                                   //LCom Version V1
                                   #statSend.tsendFct.data[#statSend.tsendFct.dataOffset] := #statSend.configTelegramV1.LComVersion;
                                   #statSend.tsendFct.data[#statSend.tsendFct.dataOffset + 1] := 16#03;
                                   #statSend.tsendFct.data[#statSend.tsendFct.dataOffset + 2] := #statSend.configTelegramV1.comMode;//ComMode
                                   #statSend.tsendFct.data[#statSend.tsendFct.dataOffset + 3] := #statSend.configTelegramV1.slidingWindow;//SlidingWindow
                                   //cycleTime
                                   #statSend.tsendFct.data[#statSend.tsendFct.dataOffset + 4] := #statSend.configTelegramV1.cycleTime.%B1;
                                   #statSend.tsendFct.data[#statSend.tsendFct.dataOffset + 5] := #statSend.configTelegramV1.cycleTime.%B0;
                                   //ackTimeOut
                                   #statSend.tsendFct.data[#statSend.tsendFct.dataOffset + 6] := #statSend.configTelegramV1.ackTimeOut.%B1;
                                   #statSend.tsendFct.data[#statSend.tsendFct.dataOffset + 7] := #statSend.configTelegramV1.ackTimeOut.%B0;
                                   //lifeSignCycle
                                   #statSend.tsendFct.data[#statSend.tsendFct.dataOffset + 8] := #statSend.configTelegramV1.lifeSignCycle.%B1;
                                   #statSend.tsendFct.data[#statSend.tsendFct.dataOffset + 9] := #statSend.configTelegramV1.lifeSignCycle.%B0;
                                   //status
                                   #statSend.tsendFct.data[#statSend.tsendFct.dataOffset + 10] := #statSend.configTelegramV1.status;
                                   //sendModeSyncTime
                                   #statSend.tsendFct.data[#statSend.tsendFct.dataOffset + 11] := #statSend.configTelegramV1.sendModeSyncTime;
                                   //maxSendDataLength
                                   #statSend.tsendFct.data[#statSend.tsendFct.dataOffset + 12] := #statSend.configTelegramV1.maxSendDataLength.%B1;
                                   #statSend.tsendFct.data[#statSend.tsendFct.dataOffset + 13] := #statSend.configTelegramV1.maxSendDataLength.%B0;
                                   //maxReceiveDataLength
                                   #statSend.tsendFct.data[#statSend.tsendFct.dataOffset + 14] := #statSend.configTelegramV1.maxReceiveDataLength.%B1;
                                   #statSend.tsendFct.data[#statSend.tsendFct.dataOffset + 15] := #statSend.configTelegramV1.maxReceiveDataLength.%B0;
                                   //calculate new offset
                                   #statSend.tsendFct.dataOffset := 16;
                               ELSE
                                   #statSend.tsendFct.data[#statSend.tsendFct.dataOffset] := #statSend.configTelegramV2.LComVersion;
                                   #statSend.tsendFct.data[#statSend.tsendFct.dataOffset + 1] := 16#03;
                                   //status
                                   #statSend.tsendFct.data[#statSend.tsendFct.dataOffset + 2] := #statSend.configTelegramV2.status;
                                   //sendModeSyncTime
                                   #statSend.tsendFct.data[#statSend.tsendFct.dataOffset + 3] := #statSend.configTelegramV2.sendModeSyncTime;
                                   //lifeSignCycle
                                   #tempDWord := TIME_TO_DWORD(#statSend.configTelegramV2.lifeSignCycle);
                                   #statSend.tsendFct.data[#statSend.tsendFct.dataOffset + 4] := #tempDWord.%B3;
                                   #statSend.tsendFct.data[#statSend.tsendFct.dataOffset + 5] := #tempDWord.%B2;
                                   #statSend.tsendFct.data[#statSend.tsendFct.dataOffset + 6] := #tempDWord.%B1;
                                   #statSend.tsendFct.data[#statSend.tsendFct.dataOffset + 7] := #tempDWord.%B0;
                                   //cycleTime
                                   #tempDWord := TIME_TO_DWORD(#statSend.configTelegramV2.cycleTime);
                                   #statSend.tsendFct.data[#statSend.tsendFct.dataOffset + 8] := #tempDWord.%B3;
                                   #statSend.tsendFct.data[#statSend.tsendFct.dataOffset + 9] := #tempDWord.%B2;
                                   #statSend.tsendFct.data[#statSend.tsendFct.dataOffset + 10] := #tempDWord.%B1;
                                   #statSend.tsendFct.data[#statSend.tsendFct.dataOffset + 11] := #tempDWord.%B0;
                                   //ackTimeOut
                                   #tempDWord := TIME_TO_DWORD(#statSend.configTelegramV2.ackTimeOut);
                                   #statSend.tsendFct.data[#statSend.tsendFct.dataOffset + 12] := #tempDWord.%B3;
                                   #statSend.tsendFct.data[#statSend.tsendFct.dataOffset + 13] := #tempDWord.%B2;
                                   #statSend.tsendFct.data[#statSend.tsendFct.dataOffset + 14] := #tempDWord.%B1;
                                   #statSend.tsendFct.data[#statSend.tsendFct.dataOffset + 15] := #tempDWord.%B0;
                                   //maxSendDataLength
                                   #statSend.tsendFct.data[#statSend.tsendFct.dataOffset + 16] := #statSend.configTelegramV2.maxSendDataLength.%B3;
                                   #statSend.tsendFct.data[#statSend.tsendFct.dataOffset + 17] := #statSend.configTelegramV2.maxSendDataLength.%B2;
                                   #statSend.tsendFct.data[#statSend.tsendFct.dataOffset + 18] := #statSend.configTelegramV2.maxSendDataLength.%B1;
                                   #statSend.tsendFct.data[#statSend.tsendFct.dataOffset + 19] := #statSend.configTelegramV2.maxSendDataLength.%B0;
                                   //maxReceiveDataLength
                                   #statSend.tsendFct.data[#statSend.tsendFct.dataOffset + 20] := #statSend.configTelegramV2.maxReceiveDataLength.%B3;
                                   #statSend.tsendFct.data[#statSend.tsendFct.dataOffset + 21] := #statSend.configTelegramV2.maxReceiveDataLength.%B2;
                                   #statSend.tsendFct.data[#statSend.tsendFct.dataOffset + 22] := #statSend.configTelegramV2.maxReceiveDataLength.%B1;
                                   #statSend.tsendFct.data[#statSend.tsendFct.dataOffset + 23] := #statSend.configTelegramV2.maxReceiveDataLength.%B0;
                                   //calculate new offset
                                   #statSend.tsendFct.dataOffset := 24;
                               END_IF;
                               #statSend.tsendFct.enable := TRUE;

                               #instLocalLifeSignCycleTimer(IN := FALSE,
                                                            PT := #diagnostics.localConfig.connection.lifeSignCycleTime);
                           ELSE
                               ;//Telegram 3 don´t need be send

                           END_IF;
                       ELSIF (NOT #diagnostics.localConfig.connection.useLComProtocol //without LCom Protocol
                           AND #statState.sender = #STATE_INACTIVE) THEN
                           #statSend.tsendFct.enable := FALSE;
                       ELSE
                           #statSend.tsendFct.enable := TRUE;

                           #instLocalLifeSignCycleTimer(IN := FALSE,
                                                        PT := #diagnostics.localConfig.connection.lifeSignCycleTime);
                       END_IF;

                       //differ between different connection types (IPv4, QDN)
                       IF (#diagnostics.localConfig.connection.connectType = #CON_TYPE_IPV4) THEN
                           #tempConnOucId := #statTconPar.ID;
                       ELSE    //#CON_TYPE_QDN
                           #tempConnOucId := #statTconParQdn.ID;
                       END_IF;

                       #instTSEND(REQ := #statSend.tsendFct.enable,
                                  LEN := #statSend.tsendFct.dataOffset,
                                  ID := #tempConnOucId,
                                  DATA := #statSend.tsendFct.data,
                                  STATUS => #statSend.tsendFct.status);

                       //16#80C4=Temporary communication error
                       IF (#statSend.tsendFct.status = 16#80C4) THEN

                           #instSendErrorTimer(IN := TRUE,
                                               PT := #MAX_TRIAL_TIME);

                           //#MAX_TRIAL_TIME is expired
                           IF #instSendErrorTimer.Q THEN
                               //Write diagnostics
                               #statDiag.bufferIndex := #statDiag.bufferIndex + 1;
                               #statDiag.buffer[#statDiag.bufferIndex].status := #ERR_SEND;
                               #statDiag.buffer[#statDiag.bufferIndex].subFunctionErrorID := #statSend.tsendFct.status;
                               #statDiag.buffer[#statDiag.bufferIndex].additionalValue1 := 0.0;
                               #statDiag.buffer[#statDiag.bufferIndex].additionalValue2 := #statSend.tsendFct.dataOffset;
                               #statDiag.buffer[#statDiag.bufferIndex].additionalValue3 := 0.0;
                               #statDiag.buffer[#statDiag.bufferIndex].additionalValue4 := T#0ms;
                               #statState.connection := #CLOSE_CONNECTION;
                               GOTO diag;
                           END_IF;
                       ELSIF (#statSend.tsendFct.status >= 16#8085) THEN
                           //#WARN_SEND
                           #statDiag.bufferIndex := #statDiag.bufferIndex + 1;
                           #statDiag.buffer[#statDiag.bufferIndex].status := #ERR_SEND;
                           #statDiag.buffer[#statDiag.bufferIndex].subFunctionErrorID := #statSend.tsendFct.status;
                           #statDiag.buffer[#statDiag.bufferIndex].additionalValue1 := 0.0;
                           #statDiag.buffer[#statDiag.bufferIndex].additionalValue2 := #statSend.tsendFct.dataOffset;
                           #statDiag.buffer[#statDiag.bufferIndex].additionalValue3 := 0.0;
                           #statDiag.buffer[#statDiag.bufferIndex].additionalValue4 := T#0ms;

                           #statState.connection := #CLOSE_CONNECTION;
                           GOTO diag;
                       END_IF;
                   END_REGION SEND_LIFESIGN

               END_REGION OPERATION

           #STATE_INACTIVE_PREPARE:
               REGION INACTIVE_PREPARE

                   #statState.connection := #STATE_INACTIVE;
                   #status := #statStatus := #STATUS_NO_CALL;
                   #statFallingEdgeEnable := FALSE;
                   #statOldEnable := FALSE;
                   #busy := FALSE;
               END_REGION INACTIVE_PREPARE

           #STATE_INIT:
               REGION INIT
                   //Reset FB Outputs
                   #connected := #statConnected := FALSE;
                   #sending := #statSending := FALSE;
                   #error := FALSE;

                   //Diagnostics purpose
                   //connection
                   #diagnostics.localConfig.connection.connectionID := #configuration.connection.connectionID;
                   #diagnostics.localConfig.connection.interfaceID := #configuration.connection.interfaceID;
                   #diagnostics.localConfig.connection.comService := #configuration.connection.comService;
                   #diagnostics.localConfig.connection.isClient := #configuration.connection.isClient;
                   #diagnostics.localConfig.connection.localPort := #configuration.connection.localPort;
                   #diagnostics.localConfig.connection.partnerPort := #configuration.connection.partnerPort;
                   #diagnostics.localConfig.connection.partnerIP := #configuration.connection.partnerIP;
                   #diagnostics.localConfig.connection.acceptUnknownPartner := #configuration.connection.acceptUnknownPartner;
                   #statActualLocalLComVersion := #HEADER_V2;
                   #diagnostics.localConfig.connection.lifeSignCycleTime := #configuration.connection.lifeSignCycleTime;
                   //-->QDN
                   #diagnostics.localConfig.connection.connectType := #configuration.connection.connectType;
                   #diagnostics.localConfig.connection.partnerQDN := #configuration.connection.partnerQDN;
                   //Sender
                   #diagnostics.localConfig.sender.cycleTime := #configuration.sender.cycleTime;
                   #diagnostics.localConfig.sender.ackTimeout := #configuration.sender.ackTimeout;
                   //TimeSync
                   #diagnostics.localConfig.timeSync.usePartnerTimestamps := #configuration.timeSync.usePartnerTimestamps;
                   #diagnostics.localConfig.timeSync.sendMode := #configuration.timeSync.sendMode;
                   #diagnostics.localConfig.timeSync.cycleTime := #configuration.timeSync.cycleTime;
                   #diagnostics.localConfig.timeSync.sendAtTimeOfDay := #configuration.timeSync.sendAtTimeOfDay;
                   //Statistics
                   #diagnostics.statistics.avgCallCycle := 0.0;
                   #diagnostics.statistics.avgReceiveMsgCycle := 0.0;
                   #diagnostics.statistics.maxReceiveMsgCycle := T#0ms;
                   #diagnostics.statistics.LComProtocolUsed := FALSE;
                   #diagnostics.statistics.activeLComVersion := 0;
                   #diagnostics.statistics.avgMsgSendingTime := 0.0;
                   #diagnostics.statistics.maxMsgSendingTime := T#0ms;
                   #diagnostics.statistics.avgMsgReceivingTime := 0.0;
                   #diagnostics.statistics.maxMsgReceivingTime := T#0ms;
                   #diagnostics.statistics.numberOfSentMessages := 0;
                   #diagnostics.statistics.numberOfReceivedMessages := 0;
                   #diagnostics.statistics.totalAckTimeouts := 0;
                   #diagnostics.statistics.totalSendCycleViolations := 0;
                   #diagnostics.statistics.totalReceiveCycleViolations := 0;
                   #diagnostics.statistics.totalReconnects := 0;

                   #statConnectAttempts := 0;

                   //Check hardware identifier of the local interface
                   IF ((#diagnostics.localConfig.connection.interfaceID >= 0) //(0...65535)
                       AND
                       (#diagnostics.localConfig.connection.interfaceID <= 65535))
                   THEN
                       //Hardware identifier of the local interface --> OK
                       #statTconPar.InterfaceId := #diagnostics.localConfig.connection.interfaceID;
                   ELSE
                       //Hardware identifier of the local interface --> NOT OK
                       #statDiag.bufferIndex := #statDiag.bufferIndex + 1;
                       #statDiag.buffer[#statDiag.bufferIndex].status := #ERR_INTERFACE_ID;
                       #statDiag.buffer[#statDiag.bufferIndex].subFunctionErrorID := 16#0000;
                       #statDiag.buffer[#statDiag.bufferIndex].additionalValue1 := UINT_TO_REAL(#diagnostics.localConfig.connection.interfaceID);//value from user
                       #statDiag.buffer[#statDiag.bufferIndex].additionalValue2 := 0.0;
                       #statDiag.buffer[#statDiag.bufferIndex].additionalValue3 := 0.0;
                       #statDiag.buffer[#statDiag.bufferIndex].additionalValue4 := T#0ms;

                       #statState.connection := #ERROR_STATE;
                       GOTO diag;
                   END_IF;

                   //Read the IP address
                   #instRDREC(REQ := TRUE,
                              ID := #configuration.connection.interfaceID,
                              INDEX := 16#8080,
                              MLEN := 0,
                              RECORD := #statSend.tsendFct.data);

                   //1st call from RDREC, to get the IP address
                   IF #instRDREC.STATUS = 16#00700100 THEN
                       ;//don´t change the #status = "STATUS_FIRST_CALL"
                   ELSE
                       //change status, that 1st call is just one time occur 
                       #status := #statStatus := #STATUS_INTERMEDIATE_CALL;
                   END_IF;

                   IF (#instRDREC.VALID = TRUE) THEN
                       //New data received and data is valid
                       #diagnostics.localConfig.connection.localIP.ADDR[1] := #statSend.tsendFct.data[28];
                       #diagnostics.localConfig.connection.localIP.ADDR[2] := #statSend.tsendFct.data[29];
                       #diagnostics.localConfig.connection.localIP.ADDR[3] := #statSend.tsendFct.data[30];
                       #diagnostics.localConfig.connection.localIP.ADDR[4] := #statSend.tsendFct.data[31];
                   ELSIF (#instRDREC.ERROR = TRUE) THEN
                       //An error occurred during the reading process
                       #diagnostics.localConfig.connection.localIP.ADDR[1] := 16#00;
                       #diagnostics.localConfig.connection.localIP.ADDR[2] := 16#00;
                       #diagnostics.localConfig.connection.localIP.ADDR[3] := 16#00;
                       #diagnostics.localConfig.connection.localIP.ADDR[4] := 16#00;
                   ELSE
                       RETURN;//The reading process is not complete yet
                   END_IF;

                   //Local port number
                   #statTconPar.LocalPort := #diagnostics.localConfig.connection.localPort;

                   //Check if send buffer is a VARIANT pointer to array of byte
                   IF ((TypeOfElements(#sendBuffer) = TypeOf(#statSend.tsendFct.data[0]))
                       AND
                       (IS_ARRAY(#sendBuffer))) THEN
                       ;//Is VARIANT pointer to array of byte
                   ELSE
                       //Write diagnostics
                       #statDiag.bufferIndex := #statDiag.bufferIndex + 1;
                       #statDiag.buffer[#statDiag.bufferIndex].status := #ERR_SEND_DATA_TYPE;
                       #statDiag.buffer[#statDiag.bufferIndex].subFunctionErrorID := 16#0000;
                       #statDiag.buffer[#statDiag.bufferIndex].additionalValue1 := 0.0;
                       #statDiag.buffer[#statDiag.bufferIndex].additionalValue2 := 0.0;
                       #statDiag.buffer[#statDiag.bufferIndex].additionalValue3 := 0.0;
                       #statDiag.buffer[#statDiag.bufferIndex].additionalValue4 := T#0ms;

                       #statState.connection := #ERROR_STATE;
                       GOTO diag;
                   END_IF;

                   //Check if receive buffer is a VARIANT pointer to array of byte
                   IF ((TypeOfElements(#receiveBuffer) = TypeOf(#statReceive.trcvFct.data[0]))
                       AND
                       (IS_ARRAY(#receiveBuffer))) THEN
                       ;//Is VARIANT pointer to array of byte
                   ELSE
                       //Write diagnostics
                       #statDiag.bufferIndex := #statDiag.bufferIndex + 1;
                       #statDiag.buffer[#statDiag.bufferIndex].status := #ERR_RECEIVE_DATA_TYPE;
                       #statDiag.buffer[#statDiag.bufferIndex].subFunctionErrorID := 16#0000;
                       #statDiag.buffer[#statDiag.bufferIndex].additionalValue1 := 0.0;
                       #statDiag.buffer[#statDiag.bufferIndex].additionalValue2 := 0.0;
                       #statDiag.buffer[#statDiag.bufferIndex].additionalValue3 := 0.0;
                       #statDiag.buffer[#statDiag.bufferIndex].additionalValue4 := T#0ms;

                       #statState.connection := #ERROR_STATE;
                       GOTO diag;
                   END_IF;

                   //Get size of user send buffer and user receive buffer in bytes
                   #diagnostics.localConfig.sizeOfSendBuffer := CountOfElements(#sendBuffer);
                   #diagnostics.localConfig.sizeOfReceiveBuffer := CountOfElements(#receiveBuffer);

                   //Check communication service: 0:UDP, 1:TCP, 2:LCOM
                   IF (#diagnostics.localConfig.connection.comService = 16#01) THEN
                       //Communication service --> transport protocol TCP
                       #statTconPar.ConnectionType := 16#0B;
                       #diagnostics.localConfig.connection.useLComProtocol := FALSE;
                   ELSIF (#diagnostics.localConfig.connection.comService = 16#02) THEN
                       //Communication service --> transport protocol TCP and LCom protocol
                       #statTconPar.ConnectionType := 16#0B;
                       #diagnostics.localConfig.connection.useLComProtocol := TRUE;
                   ELSE
                       //Communication service --> NOT OK
                       //Write diagnostics
                       #statDiag.bufferIndex := #statDiag.bufferIndex + 1;
                       #statDiag.buffer[#statDiag.bufferIndex].status := #ERR_COM_SERVICE;
                       #statDiag.buffer[#statDiag.bufferIndex].subFunctionErrorID := 16#0000;
                       #statDiag.buffer[#statDiag.bufferIndex].additionalValue1 := #diagnostics.localConfig.connection.comService;//value from operator
                       #statDiag.buffer[#statDiag.bufferIndex].additionalValue2 := 0.0;
                       #statDiag.buffer[#statDiag.bufferIndex].additionalValue3 := 0.0;
                       #statDiag.buffer[#statDiag.bufferIndex].additionalValue4 := T#0ms;

                       #statState.connection := #ERROR_STATE;
                       GOTO diag;
                   END_IF;

                   //Check unique connection identifier (16#0001...16#0FFF)
                   IF ((#diagnostics.localConfig.connection.connectionID > 0)
                       AND
                       (#diagnostics.localConfig.connection.connectionID <= 4095))
                   THEN
                       //Connection identifier -->OK
                       #statTconPar.ID := #diagnostics.localConfig.connection.connectionID;
                   ELSE
                       //Connection identifier --> NOT OK
                       //Write diagnostics
                       #statDiag.bufferIndex := #statDiag.bufferIndex + 1;
                       #statDiag.buffer[#statDiag.bufferIndex].status := #ERR_CONNECTION_ID;
                       #statDiag.buffer[#statDiag.bufferIndex].subFunctionErrorID := 16#0000;
                       #statDiag.buffer[#statDiag.bufferIndex].additionalValue1 := WORD_TO_UDINT(#diagnostics.localConfig.connection.connectionID);//value from user
                       #statDiag.buffer[#statDiag.bufferIndex].additionalValue2 := 0.0;
                       #statDiag.buffer[#statDiag.bufferIndex].additionalValue3 := 0.0;
                       #statDiag.buffer[#statDiag.bufferIndex].additionalValue4 := T#0ms;

                       #statState.connection := #ERROR_STATE;
                       GOTO diag;
                   END_IF;

                   //check connection type: 1 = IPv4, 10 = QDN
                   IF (#diagnostics.localConfig.connection.connectType = #CON_TYPE_IPV4) THEN
                       //connection type IPv4
                       ;
                   ELSIF (#diagnostics.localConfig.connection.connectType = #CON_TYPE_QDN) THEN
                       //connection type fully qualified domain name (QDN)
                       ;
                   ELSE
                       //connection type --> NOT OK
                       //write diagnostics
                       #statDiag.bufferIndex := #statDiag.bufferIndex + 1;
                       #statDiag.buffer[#statDiag.bufferIndex].status := #ERR_CONNECTION_TYPE;
                       #statDiag.buffer[#statDiag.bufferIndex].subFunctionErrorID := 16#0000;
                       #statDiag.buffer[#statDiag.bufferIndex].additionalValue1 := #diagnostics.localConfig.connection.connectType;//value from operator
                       #statDiag.buffer[#statDiag.bufferIndex].additionalValue2 := 0.0;
                       #statDiag.buffer[#statDiag.bufferIndex].additionalValue3 := 0.0;
                       #statDiag.buffer[#statDiag.bufferIndex].additionalValue4 := T#0ms;

                       #statState.connection := #ERROR_STATE;
                       GOTO diag;
                   END_IF;

                   //If client
                   IF (#diagnostics.localConfig.connection.isClient) THEN
                       //Partner port and remote address is not checked here
                       //The TCON will rise an error and return value, when the parameters (partnerPort or partnerIP) are wrong
                       //differ between different connection types (IPv4, QDN)
                       IF (#diagnostics.localConfig.connection.connectType = #CON_TYPE_IPV4) THEN
                           //remote addressing via IPv4
                           #statTconPar.RemotePort := #diagnostics.localConfig.connection.partnerPort;
                           #statTconPar.RemoteAddress := #diagnostics.localConfig.connection.partnerIP;
                       ELSE
                           //remote addressing via qualified domain name
                           #statTconParQdn.RemotePort := #diagnostics.localConfig.connection.partnerPort;
                           #statTconParQdn.RemoteQDN := #diagnostics.localConfig.connection.partnerQDN;
                           //additionally store all TCON configurations done before for QDN connection parameters
                           #statTconParQdn.ConnectionType := 16#0B;
                           #statTconParQdn.LocalPort := #diagnostics.localConfig.connection.localPort;
                           #statTconParQdn.InterfaceId := #diagnostics.localConfig.connection.interfaceID;
                           #statTconParQdn.ID := #diagnostics.localConfig.connection.connectionID;
                       END_IF;
                       //If server
                   ELSE
                       //Accept requests from all partners or only specified partner is allowed
                       IF (#diagnostics.localConfig.connection.acceptUnknownPartner) THEN
                           //Accept requests from all partners
                           //differ between different connection types (IPv4, QDN)
                           IF (#diagnostics.localConfig.connection.connectType = #CON_TYPE_IPV4) THEN
                               #statTconPar.RemoteAddress.ADDR[1] := 0;
                               #statTconPar.RemoteAddress.ADDR[2] := 0;
                               #statTconPar.RemoteAddress.ADDR[3] := 0;
                               #statTconPar.RemoteAddress.ADDR[4] := 0;
                               #statTconPar.RemotePort := 0;
                           ELSE    //#CON_TYPE_QDN
                               #statTconParQdn.RemoteQDN := '';
                               #statTconParQdn.RemotePort := 0;
                           END_IF;
                       ELSE
                           //Only specified partner is allowed
                           //differ between different connection types (IPv4, QDN)
                           IF (#diagnostics.localConfig.connection.connectType = #CON_TYPE_IPV4) THEN
                               #statTconPar.RemoteAddress := #diagnostics.localConfig.connection.partnerIP;
                               #statTconPar.RemotePort := #diagnostics.localConfig.connection.partnerPort;
                           ELSE    //#CON_TYPE_QDN
                               #statTconParQdn.RemoteQDN := #diagnostics.localConfig.connection.partnerQDN;
                               #statTconParQdn.RemotePort := #diagnostics.localConfig.connection.partnerPort;
                           END_IF;
                       END_IF;
                   END_IF;

                   //Check cycleTime
                   IF ((#diagnostics.localConfig.sender.cycleTime >= T#0ms)
                       AND
                       (#diagnostics.localConfig.sender.cycleTime <= T#+24d20h31m23s647ms))
                   THEN
                       ;//CycleTime --> OK
                   ELSE
                       //CycleTime --> NOT OK
                       #statDiag.bufferIndex := #statDiag.bufferIndex + 1;
                       #statDiag.buffer[#statDiag.bufferIndex].status := #ERR_SEND_CYCLE_TIME;
                       #statDiag.buffer[#statDiag.bufferIndex].subFunctionErrorID := 16#0000;
                       #statDiag.buffer[#statDiag.bufferIndex].additionalValue1 := 0.0;
                       #statDiag.buffer[#statDiag.bufferIndex].additionalValue2 := 0.0;
                       #statDiag.buffer[#statDiag.bufferIndex].additionalValue3 := 0.0;
                       #statDiag.buffer[#statDiag.bufferIndex].additionalValue4 := #diagnostics.localConfig.sender.cycleTime;//value from operator

                       #statState.connection := #ERROR_STATE;
                       GOTO diag;
                   END_IF;

                   //With LCom header
                   IF (#diagnostics.localConfig.connection.useLComProtocol) THEN

                       //Check lifeSignCycleTime
                       IF ((#diagnostics.localConfig.connection.lifeSignCycleTime > T#0ms) //(1ms...T#+24d20h31m23s647ms)
                           AND
                           (#diagnostics.localConfig.connection.lifeSignCycleTime <= T#+24d20h31m23s647ms))
                       THEN
                           ;//lifeSignCycleTime--> OK
                       ELSE
                           //LifeSignCycle --> NOT OK
                           #statDiag.bufferIndex := #statDiag.bufferIndex + 1;
                           #statDiag.buffer[#statDiag.bufferIndex].status := #ERR_LIFE_SIGN_CYCLE;
                           #statDiag.buffer[#statDiag.bufferIndex].subFunctionErrorID := 16#0000;
                           #statDiag.buffer[#statDiag.bufferIndex].additionalValue1 := 0.0;
                           #statDiag.buffer[#statDiag.bufferIndex].additionalValue2 := 0.0;
                           #statDiag.buffer[#statDiag.bufferIndex].additionalValue3 := 0.0;
                           #statDiag.buffer[#statDiag.bufferIndex].additionalValue4 := #diagnostics.localConfig.connection.lifeSignCycleTime;//value from operator

                           #statState.connection := #ERROR_STATE;
                           GOTO diag;
                       END_IF;

                       //Check ackTimeOut
                       IF ((#diagnostics.localConfig.sender.ackTimeout > T#0ms)
                           AND
                           (#diagnostics.localConfig.sender.ackTimeout <= T#+24d20h31m23s647ms))
                       THEN
                           ;//AckTimeOut --> OK
                       ELSE
                           //AckTimeOut --> NOT OK
                           #statDiag.bufferIndex := #statDiag.bufferIndex + 1;
                           #statDiag.buffer[#statDiag.bufferIndex].status := #ERR_ACK_TIMEOUT;
                           #statDiag.buffer[#statDiag.bufferIndex].subFunctionErrorID := 16#0000;
                           #statDiag.buffer[#statDiag.bufferIndex].additionalValue1 := 0.0;
                           #statDiag.buffer[#statDiag.bufferIndex].additionalValue2 := 0.0;
                           #statDiag.buffer[#statDiag.bufferIndex].additionalValue3 := 0.0;
                           #statDiag.buffer[#statDiag.bufferIndex].additionalValue4 := #diagnostics.localConfig.sender.ackTimeout;//value from operator

                           #statState.connection := #ERROR_STATE;
                           GOTO diag;
                       END_IF;

                       //Check timeSync
                       IF (NOT #diagnostics.localConfig.timeSync.usePartnerTimestamps) THEN

                           IF ((#diagnostics.localConfig.timeSync.sendMode >= 0)//(0...2)
                               AND
                               (#diagnostics.localConfig.timeSync.sendMode <= 2))
                           THEN
                               CASE (#diagnostics.localConfig.timeSync.sendMode) OF

                                   1: //TimeSync.cycleTime
                                       IF ((#diagnostics.localConfig.timeSync.cycleTime > T#0ms) //(1ms...T#+24d20h31m23s647ms)
                                           AND
                                           (#diagnostics.localConfig.timeSync.cycleTime <= T#+24d20h31m23s647ms))
                                       THEN
                                           ;//CycleTime --> OK
                                       ELSE
                                           //CycleTime --> Not OK
                                           #statDiag.bufferIndex := #statDiag.bufferIndex + 1;
                                           #statDiag.buffer[#statDiag.bufferIndex].status := #ERR_TIME_CYCLE_TIME;
                                           #statDiag.buffer[#statDiag.bufferIndex].subFunctionErrorID := 16#0000;
                                           #statDiag.buffer[#statDiag.bufferIndex].additionalValue1 := 0.0;
                                           #statDiag.buffer[#statDiag.bufferIndex].additionalValue2 := 0.0;
                                           #statDiag.buffer[#statDiag.bufferIndex].additionalValue3 := 0.0;
                                           #statDiag.buffer[#statDiag.bufferIndex].additionalValue4 := #diagnostics.localConfig.timeSync.cycleTime;//value from user

                                           #statState.connection := #ERROR_STATE;
                                           GOTO diag;

                                       END_IF;
                                   2://TimeSync.sendAtTimeOfDay
                                       IF ((#diagnostics.localConfig.timeSync.sendAtTimeOfDay >= TOD#00:00:00.000) //(TOD#00:00:00.000...TOD#23:59:59.999)
                                           AND
                                           #diagnostics.localConfig.timeSync.sendAtTimeOfDay <= TOD#23:59:59.999)
                                       THEN
                                           ;//SendAtTimeOfDay --> OK
                                       ELSE
                                           //SendAtTimeOfDay --> NOT OK
                                           #statDiag.bufferIndex := #statDiag.bufferIndex + 1;
                                           #statDiag.buffer[#statDiag.bufferIndex].status := #ERR_TIME_OF_DAY;
                                           #statDiag.buffer[#statDiag.bufferIndex].subFunctionErrorID := 16#0000;
                                           #statDiag.buffer[#statDiag.bufferIndex].additionalValue1 := 0.0;
                                           #statDiag.buffer[#statDiag.bufferIndex].additionalValue2 := 0.0;
                                           #statDiag.buffer[#statDiag.bufferIndex].additionalValue3 := 0.0;
                                           #statDiag.buffer[#statDiag.bufferIndex].additionalValue4 := T#0ms;

                                           #statState.connection := #ERROR_STATE;
                                           GOTO diag;
                                       END_IF;
                                   ELSE
                                       ;
                               END_CASE;
                           ELSE
                               //SendMode --> NOT OK
                               #statDiag.bufferIndex := #statDiag.bufferIndex + 1;
                               #statDiag.buffer[#statDiag.bufferIndex].status := #ERR_TIME_SYNC_MODE;
                               #statDiag.buffer[#statDiag.bufferIndex].subFunctionErrorID := 16#0000;
                               #statDiag.buffer[#statDiag.bufferIndex].additionalValue1 := #diagnostics.localConfig.timeSync.sendMode;
                               #statDiag.buffer[#statDiag.bufferIndex].additionalValue2 := 0.0;
                               #statDiag.buffer[#statDiag.bufferIndex].additionalValue3 := 0.0;
                               #statDiag.buffer[#statDiag.bufferIndex].additionalValue4 := T#0ms;

                               #statState.connection := #ERROR_STATE;
                               GOTO diag;
                           END_IF;
                       ELSE
                           //usePartnerTimeStamp

                           //Is sendMode inactive ?
                           IF #diagnostics.localConfig.timeSync.sendMode = 0 THEN
                               ;// Yes
                           ELSE
                               //SendMode --> NOT OK
                               #statDiag.bufferIndex := #statDiag.bufferIndex + 1;
                               #statDiag.buffer[#statDiag.bufferIndex].status := #ERR_TIME_SYNC_MODE;
                               #statDiag.buffer[#statDiag.bufferIndex].subFunctionErrorID := 16#0000;
                               #statDiag.buffer[#statDiag.bufferIndex].additionalValue1 := #diagnostics.localConfig.timeSync.sendMode;
                               #statDiag.buffer[#statDiag.bufferIndex].additionalValue2 := 0.0;
                               #statDiag.buffer[#statDiag.bufferIndex].additionalValue3 := 0.0;
                               #statDiag.buffer[#statDiag.bufferIndex].additionalValue4 := T#0ms;

                               #statState.connection := #ERROR_STATE;
                               GOTO diag;
                           END_IF;

                       END_IF;
                   ELSE
                       ;//No LCom Protocol is used
                   END_IF;

                   //differ between different connection types (IPv4, QDN)
                   IF (#diagnostics.localConfig.connection.connectType = #CON_TYPE_IPV4) THEN
                       //IPv4
                       #instTCON(REQ := FALSE,
                                 ID := #statTconPar.ID,
                                 CONNECT := #statTconPar);
                       //store connection ID temporary
                       #tempConnOucId := #statTconPar.ID;
                   ELSE
                       //QDN (CON_TYPE_QDN)
                       #instTCON(REQ := FALSE,
                                 ID := #statTconParQdn.ID,
                                 CONNECT := #statTconParQdn);
                       //store connection ID temporary
                       #tempConnOucId := #statTconParQdn.ID;
                   END_IF;

                   #instTSEND(REQ := FALSE,
                              ID := #tempConnOucId,
                              DATA := #statSend.tsendFct.data);

                   #instTRCV(EN_R := FALSE,
                             ID := #tempConnOucId,
                             DATA := #statReceive.trcvFct.data);

                   #instTDISCON(REQ := FALSE,
                                ID := #tempConnOucId);

                   //Passive (server), active connection establishment (client)
                   IF (#diagnostics.localConfig.connection.isClient) THEN
                       #statState.connection := #OPEN_CLIENT;
                       #statTconPar.ActiveEstablished := TRUE;
                       #statTconParQdn.ActiveEstablished := TRUE;
                   ELSE
                       #statState.connection := #OPEN_SERVER;
                       #statTconPar.ActiveEstablished := FALSE;
                       #statTconParQdn.ActiveEstablished := FALSE;
                   END_IF;
               END_REGION INIT

           #OPEN_CLIENT, #OPEN_SERVER:
               REGION OPEN_CLIENT_SERVER
                   #instTCON.STATUS := 16#0000;

                   //differ between different connection types (IPv4, QDN)
                   IF (#diagnostics.localConfig.connection.connectType = #CON_TYPE_IPV4) THEN
                       //IPv4
                       #instTCON(REQ := TRUE,
                                 CONNECT := #statTconPar,
                                 ID := #diagnostics.localConfig.connection.connectionID);
                   ELSE
                       //QDN (CON_TYPE_QDN)
                       #instTCON(REQ := TRUE,
                                 CONNECT := #statTconParQdn,
                                 ID := #diagnostics.localConfig.connection.connectionID);
                   END_IF;

                   // Error occurred
                   IF (#instTCON.ERROR) THEN

                       //Local port is being used by the system
                       IF (#instTCON.STATUS = 16#80A2 OR (#diagnostics.localConfig.connection.connectType = #CON_TYPE_IPV4 AND #statTconPar.LocalPort = 16#0)) THEN

                           #statDiag.bufferIndex := #statDiag.bufferIndex + 1;
                           #statDiag.buffer[#statDiag.bufferIndex].status := #ERR_LOCAL_PORT;
                           #statDiag.buffer[#statDiag.bufferIndex].subFunctionErrorID := #instTCON.STATUS;
                           #statDiag.buffer[#statDiag.bufferIndex].additionalValue1 := #statTconPar.LocalPort;
                           #statDiag.buffer[#statDiag.bufferIndex].additionalValue2 := 0.0;
                           #statDiag.buffer[#statDiag.bufferIndex].additionalValue3 := 0.0;
                           #statDiag.buffer[#statDiag.bufferIndex].additionalValue4 := T#0ms;

                           #statState.connection := #ERROR_STATE;
                           GOTO diag;
                           //Local port is being used by the system (in case of QDN)
                       ELSIF (#instTCON.STATUS = 16#80A2 OR (#diagnostics.localConfig.connection.connectType = #CON_TYPE_QDN AND #statTconParQdn.LocalPort = 16#0)) THEN

                           #statDiag.bufferIndex := #statDiag.bufferIndex + 1;
                           #statDiag.buffer[#statDiag.bufferIndex].status := #ERR_LOCAL_PORT;
                           #statDiag.buffer[#statDiag.bufferIndex].subFunctionErrorID := #instTCON.STATUS;
                           #statDiag.buffer[#statDiag.bufferIndex].additionalValue1 := #statTconParQdn.LocalPort;
                           #statDiag.buffer[#statDiag.bufferIndex].additionalValue2 := 0.0;
                           #statDiag.buffer[#statDiag.bufferIndex].additionalValue3 := 0.0;
                           #statDiag.buffer[#statDiag.bufferIndex].additionalValue4 := T#0ms;

                           #statState.connection := #ERROR_STATE;
                           GOTO diag;
                       ELSIF (#instTCON.STATUS = 16#80B7 OR #instTCON.STATUS = 16#80A4) THEN
                           //IP address of the remote partner is invalid
                           #statDiag.bufferIndex := #statDiag.bufferIndex + 1;
                           #statDiag.buffer[#statDiag.bufferIndex].status := #ERR_PARTNER_IP;
                           #statDiag.buffer[#statDiag.bufferIndex].subFunctionErrorID := #instTCON.STATUS;
                           #statDiag.buffer[#statDiag.bufferIndex].additionalValue1 := 0.0;
                           #statDiag.buffer[#statDiag.bufferIndex].additionalValue2 := 0.0;
                           #statDiag.buffer[#statDiag.bufferIndex].additionalValue3 := 0.0;
                           #statDiag.buffer[#statDiag.bufferIndex].additionalValue4 := T#0ms;

                           #statState.connection := #ERROR_STATE;
                           GOTO diag;
                       ELSIF (#instTCON.STATUS = 16#809B) THEN
                           //The local_device_id in the connection description does not match the CPU
                           #statDiag.bufferIndex := #statDiag.bufferIndex + 1;
                           #statDiag.buffer[#statDiag.bufferIndex].status := #ERR_INTERFACE_ID;
                           #statDiag.buffer[#statDiag.bufferIndex].subFunctionErrorID := #instTCON.STATUS;
                           #statDiag.buffer[#statDiag.bufferIndex].additionalValue1 := UINT_TO_REAL(#diagnostics.localConfig.connection.interfaceID);//value from user
                           #statDiag.buffer[#statDiag.bufferIndex].additionalValue2 := 0.0;
                           #statDiag.buffer[#statDiag.bufferIndex].additionalValue3 := 0.0;
                           #statDiag.buffer[#statDiag.bufferIndex].additionalValue4 := T#0ms;

                           #statState.connection := #ERROR_STATE;
                           GOTO diag;
                       ELSE
                           IF (#statState.connection = #OPEN_CLIENT) THEN

                               #statDiag.bufferIndex := #statDiag.bufferIndex + 1;
                               #statDiag.buffer[#statDiag.bufferIndex].status := #ERR_OPEN_CLIENT;
                               #statDiag.buffer[#statDiag.bufferIndex].subFunctionErrorID := #instTCON.STATUS;
                               #statDiag.buffer[#statDiag.bufferIndex].additionalValue1 := 0.0;
                               #statDiag.buffer[#statDiag.bufferIndex].additionalValue2 := 0.0;
                               #statDiag.buffer[#statDiag.bufferIndex].additionalValue3 := 0.0;
                               #statDiag.buffer[#statDiag.bufferIndex].additionalValue4 := T#0ms;

                               //Try reconnection after a wait time
                               #statIterator := 0;
                               #statState.connection := #STATE_WAIT;
                           ELSE
                               #statDiag.bufferIndex := #statDiag.bufferIndex + 1;
                               #statDiag.buffer[#statDiag.bufferIndex].status := #ERR_OPEN_SERVER;
                               #statDiag.buffer[#statDiag.bufferIndex].subFunctionErrorID := #instTCON.STATUS;
                               //differ between different connection types (IPv4, QDN)
                               IF (#diagnostics.localConfig.connection.connectType = #CON_TYPE_IPV4) THEN
                                   #statDiag.buffer[#statDiag.bufferIndex].additionalValue1 := #statTconPar.LocalPort;
                               ELSE    //CON_TYPE_QDN
                                   #statDiag.buffer[#statDiag.bufferIndex].additionalValue1 := #statTconParQdn.LocalPort;
                               END_IF;
                               #statDiag.buffer[#statDiag.bufferIndex].additionalValue2 := 0.0;
                               #statDiag.buffer[#statDiag.bufferIndex].additionalValue3 := 0.0;
                               #statDiag.buffer[#statDiag.bufferIndex].additionalValue4 := T#0ms;

                               //Try reconnection after a wait time
                               #statIterator := 0;
                               #statState.connection := #STATE_WAIT;
                           END_IF;
                       END_IF;
                       //Job completed without error
                   ELSIF (#instTCON.DONE) THEN

                       //Connection successfully established
                       #diagnostics.statistics.totalReconnects := #diagnostics.statistics.totalReconnects + 1;
                       #statState.connection := #OPERATION;

                       #error := FALSE;

                       //Reset all state machines
                       #statState.receiver := #READ;
                       #statState.sender := #STATE_INACTIVE;
                       #statState.comReceiver := #EXPECTED;
                       #statState.comSender := #STATE_INACTIVE;
                       //Receive
                       #statReceive.trcvFct.dataOffset := 0;
                       #statReceive.trcvFct.dataLength := 0;
                       #statReceive.trcvFct.dataLengthRest := 0;
                       #statReceive.trcvFct.dataReceived := FALSE;
                       #statReceive.tempTelegram.index := 0;
                       #statReceive.tempTelegram.telegramType := 0;
                       #statReceive.numberOfLComHeader := 0;
                       #statReceive.dataTelegram.totalMessageLength := 0;
                       #statReceive.dataTelegram.actPackageLength := 0;
                       #statReceive.dataTelegram.ackMessageOffset := 0;
                       #statReceive.dataTelegram.messageOffset := 0;
                       #statReceive.dataTelegram.ackMessageCounter := 0;
                       #statReceive.dataTelegram.messageCounter := 0;
                       #statReceive.userData.totalLength := 0;
                       #statReceive.userData.offset := 0;
                       //Send
                       #statSend.tsendFct.dataLengthRest := 0;
                       #statSend.tsendFct.dataOffset := 0;
                       #statSend.tsendFct.status := 16#0000;
                       #statSend.expectedAck.package1.offset := 0;
                       #statSend.dataTelegram.messageCounter := 0;
                       #statSend.dataTelegram.ackMessageCounter := 0;
                       #statSend.dataTelegram.messageOffset := 0;
                       #statSend.dataTelegram.ackMessageOffset := 0;
                       #statSend.dataTelegram.actPackageLength := 0;
                       #statSend.dataTelegram.totalMessageLength := 0;
                       #statSend.numberOfLComPackage := 0;
                       #statSend.userData.totalLength := 0;
                       #statSend.userData.offset := 0;
                       #statSend.userData.sendCycleViolation := FALSE;
                       #statOldSend := FALSE;

                       #diagnostics.statistics.maxMsgSendingTime := T#0ms;
                       #diagnostics.localConfig.sender.cycleTime := T#0ms;
                       #diagnostics.localConfig.sender.ackTimeout := T#0ms;

                       #diagnostics.statistics.lastTimeSync.YEAR := 2200;
                       #statCopyNBytes := 0;

                       //Reset all timer
                       #instLocalLifeSignCycleTimer(IN := FALSE,
                                                    PT := #diagnostics.localConfig.connection.lifeSignCycleTime);

                       #instPartnerLifeSignCycleTimer(IN := FALSE,
                                                      PT := (#diagnostics.partnerConfig.connnection.lifeSignCycleTime));

                       #instLocalCycleTimeTimer(IN := FALSE,
                                                PT := #diagnostics.localConfig.sender.cycleTime);

                       #instExpectedAckPackage1(IN := FALSE,
                                                PT := #diagnostics.localConfig.sender.ackTimeout);

                       #instSyncTimer(IN := FALSE,
                                      PT := T#1s);

                       #instSendErrorTimer(IN := FALSE,
                                           PT := #MAX_TRIAL_TIME);

                       #instRcvErrorTimer(IN := FALSE,
                                          PT := #MAX_TRIAL_TIME);

                       //Reset all active failures in the diagnostics buffer
                       FOR #statIterator := 0 TO #DIAG_BUFFER_UPPER_LIM BY 1 DO
                           #diagnostics.buffer[#statIterator].isActive := FALSE;
                       END_FOR;

                       //With LCom protocol
                       IF (#diagnostics.localConfig.connection.useLComProtocol = TRUE) THEN

                           IF (#statConnectAttempts MOD 2 = 0) THEN
                               //1st try LCom Version 2.0
                               #statActualLocalLComVersion := #HEADER_V2;
                               #statSend.configTelegramV2.LComVersion := #HEADER_V2;
                               #statSend.configTelegramV2.status := BOOL_TO_BYTE(#diagnostics.localConfig.timeSync.usePartnerTimestamps);
                               #statSend.configTelegramV2.sendModeSyncTime := #diagnostics.localConfig.timeSync.sendMode;
                               #statSend.configTelegramV2.lifeSignCycle := #diagnostics.localConfig.connection.lifeSignCycleTime;
                               #statSend.configTelegramV2.cycleTime := #configuration.sender.cycleTime;
                               #statSend.configTelegramV2.ackTimeOut := #configuration.sender.ackTimeout;
                               #statSend.configTelegramV2.maxSendDataLength := #diagnostics.localConfig.sizeOfSendBuffer;
                               #statSend.configTelegramV2.maxReceiveDataLength := #diagnostics.localConfig.sizeOfReceiveBuffer;

                               #statSend.dataTelegram.LComVersion := #statSend.configTelegramV2.LComVersion;
                           ELSE
                               //2nd try LCom Version 1.0
                               #statActualLocalLComVersion := #HEADER_V1;
                               #statSend.configTelegramV1.LComVersion := #HEADER_V1;
                               #statSend.configTelegramV1.comMode := 16#03;
                               #statSend.configTelegramV1.slidingWindow := 1;
                               #statSend.configTelegramV1.status := BOOL_TO_BYTE(#diagnostics.localConfig.timeSync.usePartnerTimestamps);
                               #statSend.configTelegramV1.sendModeSyncTime := #diagnostics.localConfig.timeSync.sendMode;

                               #statSend.dataTelegram.LComVersion := #statSend.configTelegramV1.LComVersion;

                               //Check max. lifeSignCycleTime
                               IF (#diagnostics.localConfig.connection.lifeSignCycleTime > T#65535ms) THEN

                                   #statDiag.bufferIndex := #statDiag.bufferIndex + 1;
                                   #statDiag.buffer[#statDiag.bufferIndex].additionalValue4 := #diagnostics.localConfig.connection.lifeSignCycleTime;
                                   #diagnostics.localConfig.connection.lifeSignCycleTime := T#65535ms;

                                   #statDiag.buffer[#statDiag.bufferIndex].status := #WARN_LIFE_SIGN_LIMITATION;
                                   #statDiag.buffer[#statDiag.bufferIndex].subFunctionErrorID := 16#0000;
                                   #statDiag.buffer[#statDiag.bufferIndex].additionalValue1 := 65535.0;
                                   #statDiag.buffer[#statDiag.bufferIndex].additionalValue2 := 0.0;
                                   #statDiag.buffer[#statDiag.bufferIndex].additionalValue3 := 0.0;
                               ELSE
                                   ;
                               END_IF;
                               #statSend.configTelegramV1.lifeSignCycle := TIME_TO_UINT(#diagnostics.localConfig.connection.lifeSignCycleTime);

                               //Check max.sizeOfSendBuffer
                               IF (#diagnostics.localConfig.sizeOfSendBuffer > 65535) THEN
                                   #diagnostics.localConfig.sizeOfSendBuffer := 65535;
                                   #statSend.configTelegramV1.maxSendDataLength := 65535;
                               ELSE
                                   #statSend.configTelegramV1.maxSendDataLength := UDINT_TO_UINT(#diagnostics.localConfig.sizeOfSendBuffer);
                               END_IF;

                               //Check max.sizeOfReceiveBuffer
                               IF (#diagnostics.localConfig.sizeOfReceiveBuffer > 65535) THEN
                                   #diagnostics.localConfig.sizeOfReceiveBuffer := 65535;
                                   #statSend.configTelegramV1.maxReceiveDataLength := 65535;
                               ELSE
                                   #statSend.configTelegramV1.maxReceiveDataLength := UDINT_TO_UINT(#diagnostics.localConfig.sizeOfReceiveBuffer);
                               END_IF;

                           END_IF;
                           //Set telegram type of data telegrams for LCom Version 1.0 and 2.0
                           #statSend.dataTelegram.telegramType := 16#0A;

                           //Start sender config directly with LCom protocol
                           #statState.cfgSender := #STATE_INIT;
                       ELSE
                           //without LCom
                           #statCompare.sender.cycleTime := #configuration.sender.cycleTime;
                           #diagnostics.localConfig.sender.cycleTime := #configuration.sender.cycleTime;

                           #diagnostics.partnerConfig.sizeOfReceiveBuffer := 0;
                           #diagnostics.partnerConfig.sizeOfSendBuffer := 0;
                           #connected := #statConnected := TRUE;
                           #statState.cfgSender := #OPERATION;

                           #statDiag.bufferIndex := #statDiag.bufferIndex + 1;
                           #statDiag.buffer[#statDiag.bufferIndex].status := #STATUS_TCP_CONNECTED;
                           #statDiag.buffer[#statDiag.bufferIndex].subFunctionErrorID := 16#0000;
                           #statDiag.buffer[#statDiag.bufferIndex].additionalValue1 := 0.0;
                           #statDiag.buffer[#statDiag.bufferIndex].additionalValue2 := 0.0;
                           #statDiag.buffer[#statDiag.bufferIndex].additionalValue3 := 0.0;
                           #statDiag.buffer[#statDiag.bufferIndex].additionalValue4 := T#0ms;
                       END_IF;
                       //TCON still in progress
                   ELSE
                       IF (#diagnostics.localConfig.connection.isClient) THEN

                           #statDiag.bufferIndex := #statDiag.bufferIndex + 1;
                           #statDiag.buffer[#statDiag.bufferIndex].status := #STATUS_CLIENT_TRY_CONNECT;
                           #statDiag.buffer[#statDiag.bufferIndex].subFunctionErrorID := 16#0000;
                           #statDiag.buffer[#statDiag.bufferIndex].additionalValue1 := 0.0;
                           #statDiag.buffer[#statDiag.bufferIndex].additionalValue2 := 0.0;
                           #statDiag.buffer[#statDiag.bufferIndex].additionalValue3 := 0.0;
                           #statDiag.buffer[#statDiag.bufferIndex].additionalValue4 := T#0ms;
                       ELSE
                           #statDiag.bufferIndex := #statDiag.bufferIndex + 1;
                           #statDiag.buffer[#statDiag.bufferIndex].status := #STATUS_SERVER_PORT_OPEN;
                           #statDiag.buffer[#statDiag.bufferIndex].subFunctionErrorID := 16#0000;
                           #statDiag.buffer[#statDiag.bufferIndex].additionalValue1 := 0.0;
                           #statDiag.buffer[#statDiag.bufferIndex].additionalValue2 := 0.0;
                           #statDiag.buffer[#statDiag.bufferIndex].additionalValue3 := 0.0;
                           #statDiag.buffer[#statDiag.bufferIndex].additionalValue4 := T#0ms;
                       END_IF;
                   END_IF;
               END_REGION OPEN_CLIENT_SERVER

           #STATE_WAIT:
               REGION WAIT
                   //Wait and then establish the connection
                   IF (#statIterator > #STATE_WAIT) THEN

                       #tempConnOucId := 0;

                       //differ between different connection types (IPv4, QDN)
                       IF (#diagnostics.localConfig.connection.connectType = #CON_TYPE_IPV4) THEN
                           //IPv4
                           #instTCON(REQ := FALSE,
                                     ID := #statTconPar.ID,
                                     CONNECT := #statTconPar);
                           //store connection ID temporary
                           #tempConnOucId := #statTconPar.ID;
                       ELSE
                           //QDN (CON_TYPE_QDN)
                           #instTCON(REQ := FALSE,
                                     ID := #statTconParQdn.ID,
                                     CONNECT := #statTconParQdn);
                           //store connection ID temporary
                           #tempConnOucId := #statTconParQdn.ID;
                       END_IF;

                       #instTSEND(REQ := FALSE,
                                  ID := #tempConnOucId,
                                  DATA := #statSend.tsendFct.data);

                       #instTRCV(EN_R := FALSE,
                                 ID := #tempConnOucId,
                                 DATA := #statReceive.trcvFct.data);

                       #instTDISCON(REQ := FALSE,
                                    ID := #tempConnOucId);

                       IF (#diagnostics.localConfig.connection.isClient) THEN
                           #statState.connection := #OPEN_CLIENT;
                           #statTconPar.ActiveEstablished := TRUE;
                           #statTconParQdn.ActiveEstablished := TRUE;
                       ELSE
                           #statState.connection := #OPEN_SERVER;
                           #statTconPar.ActiveEstablished := FALSE;
                           #statTconParQdn.ActiveEstablished := FALSE;
                       END_IF;

                   ELSE
                       #statIterator := #statIterator + 1;
                   END_IF;
               END_REGION WAIT

           #FINISH_TSEND:
               REGION FINISH_TSEND
                   IF (#statIterator > #STATE_WAIT) THEN
                       #statIterator := 0;
                       #statState.connection := #FINISH_TRCV;
                   ELSE
                       //differ between different connection types (IPv4, QDN)
                       IF (#diagnostics.localConfig.connection.connectType = #CON_TYPE_IPV4) THEN
                           #tempConnOucId := #statTconPar.ID;
                       ELSE    //CON_TYPE_QDN
                           #tempConnOucId := #statTconParQdn.ID;
                       END_IF;

                       #instTSEND(REQ := TRUE,
                                  LEN := #statSend.tsendFct.dataOffset,
                                  ID := #tempConnOucId,
                                  DATA := #statSend.tsendFct.data,
                                  STATUS => #statSend.tsendFct.status);

                       IF ((#statSend.tsendFct.status = 16#0000) OR (#instTSEND.ERROR)) THEN
                           //"TSEND" instruction is finished
                           #statState.connection := #FINISH_TRCV;
                       ELSE
                           ;//"TSEND" instruction still in process
                       END_IF;
                   END_IF;
                   #statIterator := #statIterator + 1;
               END_REGION FINISH_TSEND

           #FINISH_TRCV:
               REGION FINISH_TRCV

                   IF (#statIterator > #STATE_WAIT) THEN
                       #statState.connection := #CALL_TDISCON;
                   ELSE
                       //differ between different connection types (IPv4, QDN)
                       IF (#diagnostics.localConfig.connection.connectType = #CON_TYPE_IPV4) THEN
                           #tempConnOucId := #statTconPar.ID;
                       ELSE    //CON_TYPE_QDN
                           #tempConnOucId := #statTconParQdn.ID;
                       END_IF;

                       #instTRCV(EN_R := TRUE,
                                 ID := #tempConnOucId,
                                 LEN := 0,
                                 ADHOC := TRUE,
                                 NDR => #statReceive.trcvFct.dataReceived,
                                 RCVD_LEN => #statReceive.trcvFct.dataLength,
                                 DATA := #statReceive.trcvFct.data);

                       //Is the "TRCV" instruction still in process
                       IF (#instTRCV.ERROR OR NOT #instTRCV.BUSY) THEN
                           #statState.connection := #CALL_TDISCON;
                       ELSE
                           ;//TRCV instruction still in process
                       END_IF;
                   END_IF;
                   #statIterator := #statIterator + 1;
               END_REGION FINISH_TRCV

           #CLOSE_CONNECTION:
               REGION CLOSE_CONNECTION
                   //reset FB Outputs
                   #connected := #statConnected := FALSE;
                   #sending := #statSending := FALSE;
                   #receivedDataLength := 0;
                   #error := FALSE;

                   //Is "TSEND" instruction still in process ?
                   IF (#statSend.tsendFct.status <> 16#0000) THEN
                       //"TSEND" instruction still in process
                       #statState.connection := #FINISH_TSEND;
                       #statIterator := 0;
                   ELSE
                       ;//"TSEND" instruction is finished
                   END_IF;

                   #instTRCV(EN_R := TRUE,
                             ID := #diagnostics.localConfig.connection.connectionID,
                             LEN := 0,
                             ADHOC := TRUE,
                             NDR => #statReceive.trcvFct.dataReceived,
                             RCVD_LEN => #statReceive.trcvFct.dataLength,
                             DATA := #statReceive.trcvFct.data);

                   //Is the "TRCV" instruction still in process
                   IF (#instTRCV.ERROR OR NOT #instTRCV.BUSY) THEN
                       #statState.connection := #CALL_TDISCON;
                   ELSE
                       #statState.connection := #FINISH_TRCV;
                       #statIterator := 0;
                   END_IF;
               END_REGION CLOSE_CONNECTION

           #CALL_TDISCON:
               REGION CALL_TDISCON
                   //differ between different connection types (IPv4, QDN)
                   IF (#diagnostics.localConfig.connection.connectType = #CON_TYPE_IPV4) THEN
                       #tempConnOucId := #statTconPar.ID;
                   ELSE    //CON_TYPE_QDN
                       #tempConnOucId := #statTconParQdn.ID;
                   END_IF;

                   #instTSEND(REQ := FALSE,
                              LEN := #statSend.tsendFct.dataOffset,
                              ID := #tempConnOucId,
                              DATA := #statSend.tsendFct.data);

                   #instTRCV(EN_R := FALSE,
                             ID := #diagnostics.localConfig.connection.connectionID,
                             LEN := 0,
                             ADHOC := TRUE,
                             NDR => #statReceive.trcvFct.dataReceived,
                             RCVD_LEN => #statReceive.trcvFct.dataLength,
                             DATA := #statReceive.trcvFct.data);

                   #instTDISCON(REQ := TRUE,
                                ID := #tempConnOucId);

                   //Error occurred during processing
                   IF (#instTDISCON.ERROR) THEN

                       #statDiag.bufferIndex := #statDiag.bufferIndex + 1;
                       #statDiag.buffer[#statDiag.bufferIndex].status := #ERR_CLOSE_CONNECTION;
                       #statDiag.buffer[#statDiag.bufferIndex].subFunctionErrorID := #instTDISCON.STATUS;
                       #statDiag.buffer[#statDiag.bufferIndex].additionalValue1 := 0.0;
                       #statDiag.buffer[#statDiag.bufferIndex].additionalValue2 := 0.0;
                       #statDiag.buffer[#statDiag.bufferIndex].additionalValue3 := 0.0;
                       #statDiag.buffer[#statDiag.bufferIndex].additionalValue4 := T#0ms;

                       #statState.connection := #STATE_INACTIVE_PREPARE;

                       #instTDISCON(REQ := FALSE,
                                    ID := #tempConnOucId);

                   ELSIF (#instTDISCON.DONE) THEN

                       #instTDISCON(REQ := FALSE,
                                    ID := #tempConnOucId);
                       //Job executed without errors
                       IF (#enable AND (NOT #statFallingEdgeEnable)) THEN
                           //Reconnect automatically if not in disconnecting process
                           #statIterator := 0;
                           #statState.connection := #STATE_WAIT;
                       ELSE
                           //Reset all active failures in the diagnostics buffer
                           FOR #statIterator := 0 TO #DIAG_BUFFER_UPPER_LIM BY 1 DO
                               #diagnostics.buffer[#statIterator].isActive := FALSE;
                           END_FOR;

                           #statState.connection := #STATE_INACTIVE_PREPARE;
                       END_IF;
                       //Job is not completed yet
                   ELSE
                       ;//Wait until job is finished
                   END_IF;
               END_REGION CALL_TDISCON

           #ERROR_STATE:
               REGION ERROR
                   ;
               END_REGION ERROR
       END_CASE;
   END_REGION STATE_MACHINE

   REGION DIAGNOSTICS
       // -----------------------------------------------------------------------------------------------------------
       //Diagnostics buffer
       // -----------------------------------------------------------------------------------------------------------
   diag:
       //Diagnostics entry is in the temp. buffer
       IF (#statDiag.bufferIndex <> -1) THEN

           //Get current time
           #statRet := RD_LOC_T(#tempActTime);
           //init
           #statDiag.actualIndex := 0;

           WHILE (#statDiag.actualIndex <= #statDiag.bufferIndex) DO

               #tempUDint := 0;
               //Check if the failure is already in the buffer and still active
               FOR #statIterator := 0 TO #DIAG_BUFFER_UPPER_LIM BY 1 DO

                   IF (#diagnostics.buffer[#statIterator].isActive = TRUE) THEN

                       IF ((#statDiag.buffer[#statDiag.actualIndex].status = #WARN_SEND_CYCLE_EXPIRED)
                           AND
                           (#diagnostics.buffer[#statIterator].status = #WARN_SEND_CYCLE_EXPIRED)
                           AND
                           (#diagnostics.buffer[#statIterator].additionalValue1 = #statDiag.buffer[#statDiag.actualIndex].additionalValue1)
                           AND
                           (#diagnostics.buffer[#statIterator].additionalValue2 = #statDiag.buffer[#statDiag.actualIndex].additionalValue2)
                           AND
                           (#diagnostics.buffer[#statIterator].additionalValue3 = #statDiag.buffer[#statDiag.actualIndex].additionalValue3)) THEN
                           //Retrigger just the activation time
                           #diagnostics.buffer[#statIterator].timestamp := #tempActTime;
                           #diagnostics.buffer[#statIterator].additionalValue4 := #statDiag.buffer[#statDiag.actualIndex].additionalValue4;
                           #tempUDint := 100;
                           EXIT;
                       ELSIF ((#diagnostics.buffer[#statIterator].status = #statDiag.buffer[#statDiag.actualIndex].status)
                           AND
                           (#diagnostics.buffer[#statIterator].additionalValue1 = #statDiag.buffer[#statDiag.actualIndex].additionalValue1)
                           AND
                           (#diagnostics.buffer[#statIterator].additionalValue2 = #statDiag.buffer[#statDiag.actualIndex].additionalValue2)
                           AND
                           (#diagnostics.buffer[#statIterator].additionalValue3 = #statDiag.buffer[#statDiag.actualIndex].additionalValue3)
                           AND
                           (#diagnostics.buffer[#statIterator].additionalValue4 = #statDiag.buffer[#statDiag.actualIndex].additionalValue4)) THEN
                           //Retrigger just the activation time
                           #diagnostics.buffer[#statIterator].timestamp := #tempActTime;
                           #tempUDint := 100;
                           EXIT;
                       ELSE
                           ;//ErrorId is not in the diagnostics buffer
                       END_IF;
                   END_IF;
               END_FOR;

               IF (#tempUDint = 100) THEN
                   ;//ErrorId was already retriggered
               ELSE
                   //Check range of diagnostics ring buffer [0...DIAG_ARRAY]
                   IF ((#diagnostics.bufferIndex = 255) OR (#diagnostics.bufferIndex = #DIAG_BUFFER_UPPER_LIM)) THEN
                       #diagnostics.bufferIndex := 0;
                   ELSE
                       #diagnostics.bufferIndex := #diagnostics.bufferIndex + 1;
                   END_IF;

                   //Stored new entry in the diagnostics buffer
                   #diagnostics.buffer[#diagnostics.bufferIndex].status := #statDiag.buffer[#statDiag.actualIndex].status;
                   #diagnostics.buffer[#diagnostics.bufferIndex].timestamp := #tempActTime;
                   #diagnostics.buffer[#diagnostics.bufferIndex].isActive := TRUE;

                   #diagnostics.buffer[#diagnostics.bufferIndex].subFunctionErrorID := #statDiag.buffer[#statDiag.actualIndex].subFunctionErrorID;
                   #diagnostics.buffer[#diagnostics.bufferIndex].additionalValue1 := #statDiag.buffer[#statDiag.actualIndex].additionalValue1;
                   #diagnostics.buffer[#diagnostics.bufferIndex].additionalValue2 := #statDiag.buffer[#statDiag.actualIndex].additionalValue2;
                   #diagnostics.buffer[#diagnostics.bufferIndex].additionalValue3 := #statDiag.buffer[#statDiag.actualIndex].additionalValue3;
                   #diagnostics.buffer[#diagnostics.bufferIndex].additionalValue4 := #statDiag.buffer[#statDiag.actualIndex].additionalValue4;
               END_IF;

               IF ((#diagnostics.buffer[#diagnostics.bufferIndex].status = #STATUS_TCP_CONNECTED)
                   OR (#diagnostics.buffer[#diagnostics.bufferIndex].status = #STATUS_CONNECTED_V1)
                   OR (#diagnostics.buffer[#diagnostics.bufferIndex].status = #STATUS_CONNECTED_V2))
               THEN
                   #statConnectAttempts := 0;
                   #diagnostics.statistics.lastConnect := #tempActTime;
               END_IF;

               //Set FB status
               #status := #statStatus := #statDiag.buffer[#statDiag.actualIndex].status;

               //Check if FB.error has been set ?
               IF ((#statDiag.buffer[#statDiag.actualIndex].status >= #ERR_COM_SERVICE)//16#8200
                   AND
                   (#statDiag.buffer[#statDiag.actualIndex].status <= #ERR_WRONG_TELEGRAM_ID))//16#8614
               THEN

                   #error := TRUE;
                   #connected := #statConnected := FALSE;
                   #sending := #statSending := FALSE;
                   #dataReceived := #statDataReceived := FALSE;
                   #receivedDataLength := 0;

                   //Check if FB.busy has been set ?
                   IF ((#statDiag.buffer[#statDiag.actualIndex].status >= #ERR_OPEN_CLIENT)//16#8600
                       AND
                       (#statDiag.buffer[#statDiag.actualIndex].status <= #ERR_WRONG_TELEGRAM_ID))//16#8614
                   THEN
                       #busy := TRUE;
                   ELSE
                       #busy := FALSE;
                   END_IF;

                   EXIT;//Leave loop
               ELSE
                   ;
               END_IF;

               //Increase index
               #statDiag.actualIndex := #statDiag.actualIndex + 1;

           END_WHILE;
       ELSE
           ;//No failure
       END_IF;//End: Diagnostics buffer
   END_REGION DIAGNOSTICS
END_FUNCTION_BLOCK

FUNCTION_BLOCK "Shuttle_TCP_Comms_Shuttle2"   // FB23, SCL
{ S7_Optimized_Access := 'TRUE' }
VERSION : 0.1
// stored: AutoNumber true, IsIECCheckEnabled false, IsRetainMemResEnabled false, MemoryReserve 100, SetENOAutomatically false, UDAEnableTagReadback false
   VAR_INPUT
      Enable : Bool;
      TCP_Configuration : "LCom_typeConfig";
   END_VAR
   VAR_OUTPUT
      Connected : Bool;
      Busy : Bool;
      Status : Word;
      Error : Bool;
   END_VAR
   VAR_IN_OUT
      TCP_Diag : "LCom_typeDiagnostics";
   END_VAR
   VAR
      SendBuffer { ExternalAccessible := 'False'; ExternalVisible := 'False'; ExternalWritable := 'False'} : Array[0..1] of Byte;
      ReceiveBuffer { ExternalAccessible := 'False'; ExternalVisible := 'False'; ExternalWritable := 'False'} : Array[0..1] of Byte;
      Send : Bool;
      SendDataLength : USInt := 2;
      Sending : Bool;
   END_VAR
BEGIN
   IF "Global_Estop" THEN
       #SendBuffer[0] := 83;
       IF NOT #Send THEN
           #Send := TRUE;
       END_IF;
   ELSE
       #SendBuffer[0] := 0;
   END_IF;

   "LCom_Communication_Shuttle2_DB"(enable := #Enable,
                                    send := #Send,
                                    sendDataLength := #SendDataLength,
                                    readDataLength := 16#FFFF_FFFF,
                                    configuration := #TCP_Configuration,
                                    connected => #Connected,
                                    sending => #Sending,
                                    busy => #Busy,
                                    error => #Error,
                                    status => #Status,
                                    sendBuffer := #SendBuffer,
                                    receiveBuffer := #ReceiveBuffer,
                                    diagnostics := #TCP_Diag);

   #SendBuffer[1] := UINT_TO_BYTE("Control_DB".VTD_Control.Current_Level);

   "Control_DB".Shuttles_Position[2].Charging := "Shuttle_MQTT_DB".Shuttle_MQTT[2].Message.Shuttle_Status.Paused;

   IF #Send AND NOT #Sending THEN
       #Send := FALSE;
   END_IF;

   IF NOT #Send THEN
       "TCP_Send_Timer_DB".TON(IN := TRUE,
                               PT := T#500ms);
   END_IF;

   IF "TCP_Send_Timer_DB".Q THEN
       #Send := TRUE;
       "TCP_Send_Timer_DB".TON(IN := FALSE,
                               PT := T#0ms);
   END_IF;
END_FUNCTION_BLOCK

FUNCTION_BLOCK "Shuttle_TCP_Comms_Shuttle3"   // FB24, SCL
{ S7_Optimized_Access := 'TRUE' }
VERSION : 0.1
// stored: AutoNumber true, IsIECCheckEnabled false, IsRetainMemResEnabled false, MemoryReserve 100, SetENOAutomatically false, UDAEnableTagReadback false
   VAR_INPUT
      Enable : Bool;
      TCP_Configuration : "LCom_typeConfig";
   END_VAR
   VAR_OUTPUT
      Connected : Bool;
      Busy : Bool;
      Status : Word;
      Error : Bool;
   END_VAR
   VAR_IN_OUT
      TCP_Diag : "LCom_typeDiagnostics";
   END_VAR
   VAR
      SendBuffer { ExternalAccessible := 'False'; ExternalVisible := 'False'; ExternalWritable := 'False'} : Array[0..1] of Byte;
      ReceiveBuffer { ExternalAccessible := 'False'; ExternalVisible := 'False'; ExternalWritable := 'False'} : Array[0..1] of Byte;
      Send : Bool;
      SendDataLength : USInt := 2;
      Sending : Bool;
   END_VAR
BEGIN
   IF "Global_Estop" THEN
       #SendBuffer[0] := 83;
       IF NOT #Send THEN
           #Send := TRUE;
       END_IF;
   ELSE
       #SendBuffer[0] := 0;
   END_IF;

   "LCom_Communication_Shuttle3_DB"(enable := #Enable,
                                    send := #Send,
                                    sendDataLength := #SendDataLength,
                                    readDataLength := 16#FFFF_FFFF,
                                    configuration := #TCP_Configuration,
                                    connected => #Connected,
                                    sending => #Sending,
                                    busy => #Busy,
                                    error => #Error,
                                    status => #Status,
                                    sendBuffer := #SendBuffer,
                                    receiveBuffer := #ReceiveBuffer,
                                    diagnostics := #TCP_Diag);

   #SendBuffer[1] := UINT_TO_BYTE("Control_DB".VTD_Control.Current_Level);

   "Control_DB".Shuttles_Position[3].Charging := "Shuttle_MQTT_DB".Shuttle_MQTT[3].Message.Shuttle_Status.Paused;

   IF #Send AND NOT #Sending THEN
       #Send := FALSE;
   END_IF;

   IF NOT #Send THEN
       "TCP_Send_Timer_DB".TON(IN := TRUE,
                               PT := T#500ms);
   END_IF;

   IF "TCP_Send_Timer_DB".Q THEN
       #Send := TRUE;
       "TCP_Send_Timer_DB".TON(IN := FALSE,
                               PT := T#0ms);
   END_IF;
END_FUNCTION_BLOCK

FUNCTION "OUTPUTS" : Void   // FC5, SCL
{ S7_Optimized_Access := 'TRUE' }
VERSION : 0.1
// stored: AutoNumber true, IsIECCheckEnabled false, SetENOAutomatically false, UDAEnableTagReadback false
BEGIN

   // Let's do it for each Shuttle 
   //IF destinationid = position id = id charger (*Setpoint in the HMI reggarding to the charger position*)
   //     2000 = 2000 = 2000 // Example 1 Shuttle on charger positio => Charger on
   //     2000 = 1900 = 2000 // Example 2 Shuttle in other position => Charger off
   //     1000 = 2000 = 2000 // Example 3 Shuttle in charger position but received an order to move to other position => Charger off
   // Enable the charger (Variable) = TRUE;
   //ELSE  
     // Disable the charger
     // Enable the charger (Variable) = FALSE;
   //END_IF;


   IF "FirstScan" THEN
       "Charger Panel" := TRUE;
   END_IF;

   "Charger Panel" := "Charger";

   "Pick Station light" := "Control_DB".Pick_Station.PushButtonLight;
END_FUNCTION

FUNCTION_BLOCK "Order_Table_FB_Carousel"   // FB32, SCL
{ S7_Optimized_Access := 'TRUE' }
VERSION : 0.1
// stored: AutoNumber true, IsIECCheckEnabled false, IsRetainMemResEnabled false, MemoryReserve 100, SetENOAutomatically false, UDAEnableTagReadback false
   VAR_INPUT
      System_Selected { ExternalWritable := 'False'} : Bool;
      AutoMan_Switch : Bool;   // Auto/Man Switch on CPU Panel - 1 = Auto, 0 = Manual
      CurrentTime { ExternalWritable := 'False'} : String;
      CurrentDTL : DTL;
      Watchdog : "Watchdog_Settings_UDT";
   END_VAR
   VAR_IN_OUT
      Cnv_Entry : "Inbound_Cnv_Control_UDT";
      Cnv_PopUp_1 : "PopUp_Cnv_Control";
      WeighingStation : "Stations_DB_UDT";
      ProfileStation : "Stations_DB_UDT";
      Cnv_PopUp_2 : "PopUp_Cnv_Control";
      Cnv_PopUp_3 : "PopUp_Cnv_Control";
      Cnv_PopUp_4 : "PopUp_Cnv_Control";
      Cnv_Exit : "Outbound_Cnv_Control";
      System : "System_UDT";
      Control_OPC_Ua : "WMS_OPC_UA";
   END_VAR
   VAR
      RTR_ITP1_CurrentOrder : UDInt;
      RTR_P1P2_CurrentOrder : UDInt;
      RTR_P3P4_CurrentOrder : UDInt;
      RTR_P4TO_CurrentOrder : UDInt;
      Roller_To_Roller_CurrentOrder : UDInt;
      Chain_To_Chain_CurrentOrder : UDInt;
      Pop4_To_PickSt_CurrentOrder : UDInt;
      PickSt_To_Pop1_CurrentOrder : UDInt;
      WeighingStation_CurrentOrder { ExternalWritable := 'False'} : UDInt := 0;
      ProfileStation_CurrentOrder { ExternalWritable := 'False'} : UDInt := 0;
      Roller_To_RollerDoneRTrig : R_TRIG;
      RTR_ITP1DoneRTrig { S7_SetPoint := 'True'} : R_TRIG;
      RTR_P1P2DoneRTrig { S7_SetPoint := 'True'} : R_TRIG;
      RTR_P3P4DoneRTrig { S7_SetPoint := 'True'} : R_TRIG;
      RTR_P4TODoneRTrig { S7_SetPoint := 'True'} : R_TRIG;
      Chain_To_ChainDoneRTrig : R_TRIG;
      Pop4_To_PickSt_DoneRTrig { S7_SetPoint := 'True'} : R_TRIG;
      PickSt_To_Pop1_DoneRTrig { S7_SetPoint := 'True'} : R_TRIG;
      WeighingStationDoneRTrig { ExternalWritable := 'False'} : R_TRIG;
      ProfileStationDoneRTrig { ExternalWritable := 'False'} : R_TRIG;
      PalletRefused_1_RTig { ExternalWritable := 'False'} : R_TRIG;
      ErrorRTrig { ExternalWritable := 'False'} : R_TRIG;
      CancelRTrig { ExternalWritable := 'False'} : R_TRIG;
      PauseRTrig { ExternalWritable := 'False'} : R_TRIG;
      ResumeRTrig { ExternalWritable := 'False'} : R_TRIG;
      Clear_Store : R_TRIG;
      Clear_Retrieve : R_TRIG;
      Canceling : Bool;
      RTR_ITP1_WatchdogTimer : TON_TIME;
      RTR_P1P2_WatchdogTimer : TON_TIME;
      RTR_P3P4_WatchdogTimer : TON_TIME;
      RTR_P4TO_WatchdogTimer : TON_TIME;
      Roller_To_Roller_WatchdogTimer { S7_SetPoint := 'True'} : TON_TIME;
      Chain_To_Chain_WatchdogTimer { S7_SetPoint := 'True'} : TON_TIME;
      Pop4_To_PickWatchdogTimer { S7_SetPoint := 'True'} : TON_TIME;
      PickSt_To_Pop1WatchdogTimer : TON_TIME;
      WeighingStation_WatchdogTimer : TON_TIME;
      ProfileStation_WatchdogTimer : TON_TIME;
      Roller_To_Roller_WatchdogStart { S7_SetPoint := 'True'} : Bool;
      RTR_ITP1_WatchdogStart : Bool;
      RTR_P1P2_WatchdogStart : Bool;
      RTR_P3P4_WatchdogStart : Bool;
      RTR_P4TO_WatchdogStart : Bool;
      Chain_To_Chain_WatchdogStart : Bool;
      Pop4_To_PickWatchdogStart : Bool;
      PickSt_To_Pop1WatchdogStart : Bool;
      WeighingStation_WatchdogStart : Bool;
      ProfileStation_WatchdogStart : Bool;
      dummy : Int;
      dummy_1 : Bool;
      dummy_3 : Bool;
   END_VAR
   VAR_TEMP
      i : DInt;
      n : DInt;
      EmptyOrder : "OrderTable_UDT";
      MaxRunningOrderNo : UInt;
   END_VAR
   VAR CONSTANT
      RTR_ITOP1 : String := 'RTR ITP1';
      RTR_P1_TO_P2 : String := 'RTR P1P2';
      RTR_P3_TO_P4 : String := 'RTR P3P4';
      RTR_P4TO : String := 'RTR P4TO';
      ROLLER_TO_ROLLER_DEVICE : String := 'Roller to Roller';
      CHAIN_TO_CHAIN_DEVICE : String := 'Chain to Chain';
      POP4_TO_PICK_DEVICE : String := 'Pop4 to Pick';
      PICK_TO_POP1_DEVICE : String := 'Pick to Pop1';
      WEIGH_STATION_DEVICE : String := 'Weigh Station';
      PROFILE_STATION_DEVICE : String := 'Profile Station';
      RUNNING_STATUS : String := 'Running';
      COMPLETED_STATUS : String := 'Completed';
      QUEUED_STATUS : String := 'Queued';
      PALLET_REFUSED_STATUS : String := 'Pallet Refused';
      ERROR_STATUS : String := 'Error';
      CANCELED_STATUS : String := 'Canceled';
      PAUSED_STATUS : String := 'Paused';
      ORDER_REFUSED : String := 'Refused';
      ERROR_CANCELED_STATUS : String := 'Error\Cancel';
   END_VAR
BEGIN

   // Converts the task type for strings 
   IF #System.OrderTable[1].OPC_Control.Task_Type = 6
           AND #System.OrderTable[1].OPC_Control.Destination_Location = 140001 THEN // Roller to Roller - Outbound Conveyor final destination
           #System.OrderTable[1].Device := 'RTR P4TO';
   ELSIF #System.OrderTable[1].OPC_Control.Task_Type = 6
           AND #System.OrderTable[1].OPC_Control.Destination_Location = 180001  THEN // Roller to Roller - Pop conveyor 4 - final destination
           #System.OrderTable[1].Device := 'RTR P3P4';
       ELSIF #System.OrderTable[1].OPC_Control.Task_Type = 6
           AND #System.OrderTable[1].OPC_Control.Destination_Location = 160001  THEN // Roller to Roller - Pop conveyor 4 - final destination
           #System.OrderTable[1].Device := 'RTR P1P2';
       ELSIF #System.OrderTable[1].OPC_Control.Destination_Location = 150001 AND (#System.OrderTable[1].OPC_Control.Task_Type = 16 OR #System.OrderTable[1].OPC_Control.Task_Type = 6) THEN //Roller TO Roller + Barcode scanner
       #System.OrderTable[1].Device := 'RTR ITP1';
   ELSIF #System.OrderTable[1].OPC_Control.Task_Type = 14 THEN //Roller TO Roller + Profile Station
       #System.OrderTable[1].Device := 'RTR P1P2';
   ELSIF #System.OrderTable[1].OPC_Control.Task_Type = 7 THEN
       #System.OrderTable[1].Device := 'Chain to Chain';
   ELSIF #System.OrderTable[1].OPC_Control.Task_Type = 8 THEN
       #System.OrderTable[1].Device := 'Pop4 to Pick';
   ELSIF #System.OrderTable[1].OPC_Control.Task_Type = 9 THEN
       #System.OrderTable[1].Device := 'Pick to Pop1' ;
   ELSIF #System.OrderTable[1].OPC_Control.Task_Type = 10 THEN
       #System.OrderTable[1].Device := 'Weigh Station';
   // ELSIF #System.OrderTable[1].OPC_Control.Task_Type = 14 THEN
   //     #System.OrderTable[1].Device := 'Profile Station';
   ELSE
       #System.OrderTable[1].Device := '';
   END_IF;


   REGION #New Order was Sent
       IF #System.OrderSent THEN
           //Count orders in Step Table
           FOR #i := 0 TO 20 DO
               IF #System.StepTable[#i].OrderNo <> 0
                   AND #System.StepTable[#i].StepNo <> 0
                   AND #System.StepTable[#i].PlaceTime <> ''
                   //AND #System.StepTable[#i].Device <> ''
                   AND #System.StepTable[#i].Status = #QUEUED_STATUS
               THEN
                   #n += 1;
               ELSE
                   EXIT;
               END_IF;
           END_FOR;

           IF #n > 0 THEN
               //shift order table down by Order number rows
               FOR #i := 99 TO (#n + 1) BY -1 DO
                   #System.OrderTable[#i] := #System.OrderTable[#i - #n];
               END_FOR;
               //copy data from step table to order table
               FOR #i := 0 TO #n DO
                   #System.OrderTable[#n - #i (*+ 1*)] := #System.StepTable[#i];
               END_FOR;
               //clean step table
               FOR #i := 0(*1*) TO 20 DO
                   #System.StepTable[#i] := #EmptyOrder;
               END_FOR;
               #System.CurrentOrder += #n;


               // // Transfer Pallet Roller to Roller - 

               // IF #Roller_To_Roller_CurrentOrder <> 0 THEN
               //     #Roller_To_Roller_CurrentOrder += #n;
               // END_IF;


               // Transfer Pallet Roller to Roller - Inbound to PP1

               IF #RTR_ITP1_CurrentOrder <> 0 THEN
                   #RTR_ITP1_CurrentOrder += #n;
               END_IF;

               // Transfer Pallet Roller to Roller - PP1 to PP2

               IF #RTR_P1P2_CurrentOrder <> 0 THEN
                   #RTR_P1P2_CurrentOrder += #n;
               END_IF;

               // Transfer Pallet Roller TO Roller - PP3 TO PP4

               IF #RTR_P3P4_CurrentOrder <> 0 THEN
                   #RTR_P3P4_CurrentOrder += #n;
               END_IF;


               // Transfer Pallet Roller TO Roller - PP4 TO OUTBOUND

               IF #RTR_P4TO_CurrentOrder <> 0 THEN
                   #RTR_P4TO_CurrentOrder += #n;
               END_IF;


               // Transfer Pallet Chain to Chain
               IF #Chain_To_Chain_CurrentOrder <> 0 THEN
                   #Chain_To_Chain_CurrentOrder += #n;
               END_IF;

               // Transfer TO pick station (From Pop Conveyor 4)
               IF #Pop4_To_PickSt_CurrentOrder <> 0 THEN
                   #Pop4_To_PickSt_CurrentOrder += #n;
               END_IF;

               // Transfer from Pick station (To Pop Conveyor 1)
               IF #PickSt_To_Pop1_CurrentOrder <> 0 THEN
                   #PickSt_To_Pop1_CurrentOrder += #n;
               END_IF;


               //Weigh Station
               IF #WeighingStation_CurrentOrder <> 0 THEN
                   #WeighingStation_CurrentOrder += #n;
               END_IF;

               //Profile Station
               IF #ProfileStation_CurrentOrder <> 0 THEN
                   #ProfileStation_CurrentOrder += #n;
               END_IF;


           END_IF;
            #System.OrderSent := FALSE;
       END_IF;
   END_REGION

   REGION Auto/Man Mode
       //Enable Devices in Auto/Man Mode
       IF #System.Auto_Man THEN
         //  #Cnv_Entry.Mode := #Cnv_PopUp_1.Mode:= #WeighingStation.Mode := #ProfileStation.Mode :=
          // #Cnv_PopUp_2.Mode := #Cnv_PopUp_3.Mode := #Cnv_PopUp_4.Mode := #Cnv_Exit.Mode := 3;// Auto Mode

           #Cnv_Entry.Instruction.Enable := #Cnv_PopUp_1.Instruction.Enable := #WeighingStation.Enable :=
           #ProfileStation.Enable := #Cnv_PopUp_2.Instruction.Enable := #Cnv_PopUp_3.Enabled := #Cnv_PopUp_4.Instruction.Enable :=
           #Cnv_Exit.Instruction.Enable := TRUE; // := Not System.Error

       ELSE //Disable Devices in Auto/Man Mode
          // #Cnv_Entry.Mode := #Cnv_PopUp_1.Mode := #WeighingStation.Mode := #ProfileStation.Mode :=
         //  #Cnv_PopUp_2.Mode := #Cnv_PopUp_3.Mode := #Cnv_PopUp_4.Mode := #Cnv_Exit.Mode:= 0;
           #Cnv_Entry.Instruction.Enable := #Cnv_PopUp_1.Instruction.Enable := #WeighingStation.Enable :=
           #ProfileStation.Enable := #Cnv_PopUp_2.Instruction.Enable := #Cnv_PopUp_3.Enabled := #Cnv_PopUp_4.Instruction.Enable :=
           #Cnv_Exit.Instruction.Enable := FALSE;
       END_IF;
   END_REGION

   REGION Roller TO Roller - Carousel Conveyors - Inbound to PP1 - With Barcode
   //Roller conveyors
   IF #System.OrderTable[1].StepNo <> 0
       AND #System.OrderTable[1].Device = #RTR_ITOP1
       AND #System.OrderTable[1].Status = #QUEUED_STATUS
       AND "OPC_UA_Control_FB_DB".State_Carrousel_ITP1 = 0
       AND NOT #System.Error
       AND NOT #Canceling

   THEN
       #RTR_ITP1_CurrentOrder := 1;
   END_IF;
   IF #System.OrderTable[#RTR_ITP1_CurrentOrder].StepNo <> 0
       AND #System.OrderTable[#RTR_ITP1_CurrentOrder].Device = #RTR_ITOP1
       AND #System.OrderTable[#RTR_ITP1_CurrentOrder].Status = #QUEUED_STATUS
       AND "OPC_UA_Control_FB_DB".State_Carrousel_ITP1 = 0
       AND NOT #System.Error
       AND NOT #Canceling

   THEN
       //OPC Commands to Move Pallets - Carousel Conveyors
       // WCS => Order Table => OPC Ua Control Table

       IF #System.OrderTable[1].OPC_Control.Task_Type = 16 THEN // Barcode Scanner - INB TO P1
           "Control_DB"."InBarcode_Station".Start := TRUE;
       ELSE
           "Control_DB"."InBarcode_Station".Start := FALSE;
       END_IF;

       "Control_DB"."Carrousel_Order Table".Task_Data_Available := TRUE;//#System.OrderTable[#Roller_To_Roller_CurrentOrder].OPC_Control.Task_Data_Available; // Send the Task Data Available from WCS 
       "Control_DB"."Carrousel_Order Table".Task_Type := #System.OrderTable[#RTR_ITP1_CurrentOrder].OPC_Control.Task_Type; //  Send the Task Type - Roller to Roller Conveyor = Task Type = 6
       "Control_DB"."Carrousel_Order Table".Task_ID := #System.OrderTable[#RTR_ITP1_CurrentOrder].OPC_Control.Task_ID; // Send the Task ID number;
       "Control_DB"."Carrousel_Order Table".Task_Metadata := #System.OrderTable[#RTR_ITP1_CurrentOrder].OPC_Control.Task_Metadata; // Send the Task Metadata Unique identifier
       "Control_DB"."Carrousel_Order Table".Source_Location := #System.OrderTable[#RTR_ITP1_CurrentOrder].OPC_Control.Source_Location; // Send the Source Location from the Conveyor
       "Control_DB"."Carrousel_Order Table".Destination_Location := #System.OrderTable[#RTR_ITP1_CurrentOrder].OPC_Control.Destination_Location; // Send the Destination Location to the Conveyor;
       #Roller_To_Roller_WatchdogStart := true;


   END_IF;

   //RUNNING
   IF "OPC_UA_Control_FB_DB".State_Carrousel_ITP1 > 0 AND "OPC_UA_Control_FB_DB".State_Carrousel_ITP1 < 400  AND #System.Auto_Man THEN
       #System.OrderTable[#RTR_ITP1_CurrentOrder].Status := #RUNNING_STATUS;
   END_IF;

   //Cancel order
   IF #Canceling AND NOT (#Cnv_Entry.Running OR #Cnv_PopUp_1.Running) AND #RTR_ITP1_CurrentOrder <> 0
   THEN
       #System.OrderTable[#RTR_ITP1_CurrentOrder].Status := #CANCELED_STATUS;
       #System.OrderTable[#RTR_ITP1_CurrentOrder].CompleteTime := #CurrentTime;
       #RTR_ITP1_CurrentOrder := 0;


       "Control_DB".InBarcode_Station.Start := FALSE;
       "Control_DB"."Carrousel_Order Table".Task_Data_Available := FALSE; // Send the Task Data Available from WCS 
       "Control_DB"."Carrousel_Order Table".Task_Type := 0; //  Send the Task Type - Roller to Roller Conveyor = Task Type = 6
       "Control_DB"."Carrousel_Order Table".Task_ID := 0; // Send the Task ID number;
       "Control_DB"."Carrousel_Order Table".Task_Metadata := ''; // Send the Task Metadata Unique identifier
       "Control_DB"."Carrousel_Order Table".Source_Location := 0; // Send the Source Location from the Conveyor
       "Control_DB"."Carrousel_Order Table".Destination_Location := 0; // Send the Destination Location to the Conveyor;

   END_IF;

   //Error
   IF (#Cnv_Entry.Error OR #Cnv_PopUp_1.Error) THEN
       //#Cnv_Entry.Instruction.Execute := FALSE;

       "Control_DB".InBarcode_Station.Start := FALSE;
       "Control_DB"."Carrousel_Order Table".Task_Data_Available := FALSE; // Send the Task Data Available from WCS 
       "Control_DB"."Carrousel_Order Table".Task_Type := 0; //  Send the Task Type - Roller to Roller Conveyor = Task Type = 6
       "Control_DB"."Carrousel_Order Table".Task_ID := 0; // Send the Task ID number;
       "Control_DB"."Carrousel_Order Table".Task_Metadata := ''; // Send the Task Metadata Unique identifier
       "Control_DB"."Carrousel_Order Table".Source_Location := 0; // Send the Source Location from the Conveyor
       "Control_DB"."Carrousel_Order Table".Destination_Location := 0; // Send the Destination Location to the Conveyor;
       #System.OrderTable[#RTR_ITP1_CurrentOrder].ErrorID := (#Cnv_Entry.Cnv_Errors.Error_Word_4
       OR #Cnv_PopUp_1.Cnv_Errors.Error_Word_1
       );

   END_IF;

   //MOVEMENT FINALIZED
   #RTR_ITP1DoneRTrig(CLK := "Control_DB".Movement_Completed.RTR_ITP1);
   IF #RTR_ITP1DoneRTrig.Q THEN
       "Control_DB".Movement_Completed.RTR_ITP1 := FALSE;

       "Control_DB".InBarcode_Station.Start := FALSE;
       "Control_DB"."Carrousel_Order Table".Task_Data_Available := FALSE; // Send the Task Data Available from WCS 
       "Control_DB"."Carrousel_Order Table".Task_Type := 0; //  Send the Task Type - Roller to Roller Conveyor = Task Type = 6
       "Control_DB"."Carrousel_Order Table".Task_ID := 0; // Send the Task ID number;
       "Control_DB"."Carrousel_Order Table".Task_Metadata := ''; // Send the Task Metadata Unique identifier
       "Control_DB"."Carrousel_Order Table".Source_Location := 0; // Send the Source Location from the Conveyor
       "Control_DB"."Carrousel_Order Table".Destination_Location := 0; // Send the Destination Location to the Conveyor;

       #RTR_ITP1_WatchdogStart := FALSE;
       #System.OrderTable[#RTR_ITP1_CurrentOrder].Status := #COMPLETED_STATUS;
       #System.OrderTable[#RTR_ITP1_CurrentOrder].CompleteTime := #CurrentTime;
       #RTR_ITP1_CurrentOrder := 0;
   END_IF;
   END_REGION

   REGION Roller TO Roller - Carousel Conveyors - PP1 to PP2 - With Profile Station
       //Roller conveyors
       IF #System.OrderTable[1].StepNo <> 0
           AND #System.OrderTable[1].Device = #RTR_P1_TO_P2
           AND #System.OrderTable[1].Status = #QUEUED_STATUS
           AND NOT (#Cnv_PopUp_1.Running OR #Cnv_PopUp_2.Running)
           AND NOT #System.Error
           AND NOT #Canceling

       THEN
           #RTR_P1P2_CurrentOrder := 1;
       END_IF;
       IF #System.OrderTable[#RTR_P1P2_CurrentOrder].StepNo <> 0
           AND #System.OrderTable[#RTR_P1P2_CurrentOrder].Device = #RTR_P1_TO_P2
           AND #System.OrderTable[#RTR_P1P2_CurrentOrder].Status = #QUEUED_STATUS
           AND NOT (#Cnv_PopUp_1.Running OR #Cnv_PopUp_2.Running)
           AND NOT #System.Error
           AND NOT #Canceling

       THEN
           //OPC Commands to Move Pallets - Carousel Conveyors
           // WCS => Order Table => OPC Ua Control Table

           IF #System.OrderTable[1].OPC_Control.Task_Type = 14 THEN // Profile Station - P1 TO P2
               "Control_DB"."Profiling Station".Start := TRUE;
           ELSE
               "Control_DB"."Profiling Station".Start := FALSE;
           END_IF;

